(* Logix 5000 project; controller R400_500_XLS vendor 1 type 14 code 216 rev 31.11; software revision 31.01; part 27 of 32 *)
(* tags used below, declared in another part *)
   Abort1 : DINT;   // Not Used
   Alarm : SINT;   // Wait 3 seconds
   AlarmAcked : BOOL;   // Alarm has been acked
   Ashutdown : SINT;   // Not Used
   bAlrm : BOOL[64];
   Change_PrintPtr_Value : BOOL;
   CHEMICAL_COND_MAX_TIME : DINT;   // Timeout for the conductivity based chemical injection
   CHEMICAL_PUMP_OFF_TIME : DINT[4];
   CHEMICAL_PUMP_ON_TIME : DINT[4];
   CycExcBuffer : UDT_CYCLE;
   CycleSequence : UDT_CYCLE_SEQUENCE;
   CycleTime : DINT[11];   // Last cycle time saved in seconds
   DRYING : DINT;   // Drying id number
   FC23_BaseConductivity : REAL;   // Base conductivity of the water prior to the injection
   FC23_ChemicalPumpIndex : DINT;   // Chemical pump index
   FC23_CompensatedSetPoint : REAL;   // Injection compensated chemical conductivity
   FC23_FinalConductivity : REAL;   // Final value of the chemical conductivity
   FC23_OffsetSetPoint : REAL;   // Set point before enabling the on/off sequence
   FC23_ONS : SINT;
   FC23_StartSignal : BOOL;   // Conductivity based chemical injection
   FC23_WashIndex : DINT;   // Current index of the wash treatment
   FINALRINSE_1 : DINT;   // Final rinse 1 id number
   Inj_Cond : SINT;   // Conductivity injection based steps
   Inj_Cond_Tran : SINT;   // Conductivity injection based transitions
   InjMan : SINT;
   M : DINT[5];   // Memory Bits
   New_Value : SINT;
   ONS_FC24 : SINT;
   ONS_FC37 : DINT;
   ONS_FC64 : DINT;
   OPR_16_TreatPrint_Ptr : DINT;
   PREWASH_1 : DINT;   // Pre-wash 1 id number
   PREWASH_2 : DINT;   // Pre-wash 2 id number
   PREWASH_3 : DINT;   // Pre-wash 3 id number
   PREWASH_4 : DINT;   // Pre-wash 4 id number
   Print_Data : BOOL;   // Print Treatment data
   Print_Speed_Water : BOOL;
   Print_TreatEnd_Start_Data : BOOL;   // 2nd treatment of the cycle is started, pirnt Treatment Completed and Treatment data
   Print_TreatStart_Data : BOOL;   // Cycle is started Print start time and treatment data of the first treatment of the cycle
   printTreatString : STRING[85];   // Treatment String
   PWR_PrintBuffer : UDT_WASH;
   rIn_WSH61 : REAL;
   RINSE_1 : DINT;   // Rinse 1 id number
   RINSE_2 : DINT;   // Rinse 2 id number
   RINSE_3 : DINT;   // Rinse 3 id number
   RINSE_4 : DINT;   // Rinse 4 id number
   Run : DINT;
   sCRLF : STRING;
   SET_POINT_FRACTION : REAL[4];
   sFll_Zero : STRING[20];
   SMART_MODE_DRYING_HEATCOOL_SEC : DINT;   // Heating and cooling time constant for the smart mode drying (sec.)
   sOut_WSH61 : STRING;
   sPrntArray : STRING[300];   // Printer String Array
   SRE3_Serial_Number : STRING;   // Serial number
   StartPump3 : BOOL;   // Main Pump running
   String : STRING[50];   // String
   String_Temp : STRING;
   Tmr : TIMER[107];
   TreatmentPrint_Ptr : SINT;
   Trt_Drying : SINT;
   Trt_Wsh : DINT;
   VENTING : DINT;   // Venting id number
   WASH_1 : DINT;   // Wash 1 id number
   WASH_2 : DINT;   // Wash 2 id number
   WASH_3 : DINT;   // Wash 3 id number
   WASH_4 : DINT;   // Wash 4 id number
   WASH_5 : DINT;   // Wash 5 id number
   WSH36_CycleTimePercentage : DINT;
   WSH36_SecondsRemaining : DINT;
   WSH36_TotalMinutesRemaining : DINT;
   WSH36_TotalSecondsRemaining : DINT;
   WSH41_Start_signal : BOOL;   // Start cycle signal One shot rising edge
   WSH56_TreatmentInfo : BOOL;   // Treatment information for the conductivity injection
   Zero_Value : SINT;
   ChemCond : REAL;
   ChemicalName : STRING[9];   // Used by HMI
   COOLING_PHASE_TIME : DINT;   // Time of the cooling phase when time based drying
   CyclePtr : DINT;   // Cycle Pointeur
   I_Chm_1_Lvl_Sw : BOOL;   // Chemical Pump #1 level switch
   I_Chm_2_Lvl_Sw : BOOL;   // Chemical Pump #2 level switch
   I_Chm_3_Lvl_Sw : BOOL;   // Chemical Pump #3 level switch
   I_Chm_4_Lvl_Sw : BOOL;   // Chemical Pump #4 level switch
   Load : Doors;
   PrintChemCondValue : REAL;
   printID : STRING[6];
   PrintIndex : DINT;
   rSCADACompensatedSetPoint : REAL;
   Screen_Ctrl : DINT;   // PLC Screen Request
   sTime : STRING;   // String current time
   SumpTemp : REAL;   // Sump temperature in °C
   TempUnit : BOOL;   // Temperature Units 0= Celcius 1 = Farhenheit
   Tpb : DINT[11];
   TreatmentPtr : DINT;
   Unit : Hrdwre;   // Unit Configuration
(* MainProgram, continued *)

ROUTINE WSH_33_MANUAL_INJECTION   (* ladder *)
// This routine manages the manual  chemical injection
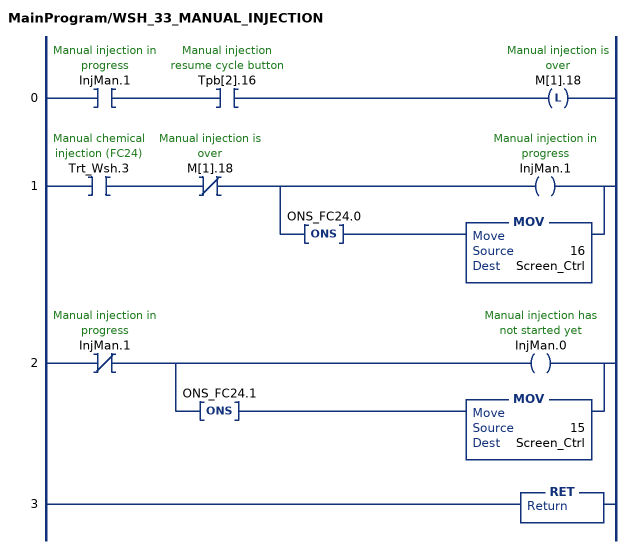
   0: XIC(InjMan.1)XIC(Tpb[2].16)OTL(M[1].18);
   1: XIC(Trt_Wsh.3)XIO(M[1].18)[OTE(InjMan.1) ,ONS(ONS_FC24.0) MOV(16,Screen_Ctrl) ];
   2: XIO(InjMan.1)[OTE(InjMan.0) ,ONS(ONS_FC24.1) MOV(15,Screen_Ctrl) ];
   3: RET();
END_ROUTINE

ROUTINE WSH_34_CONDUCTIVITY_INJECTION   (* ladder *)
// This routine manages the time based chemical injection
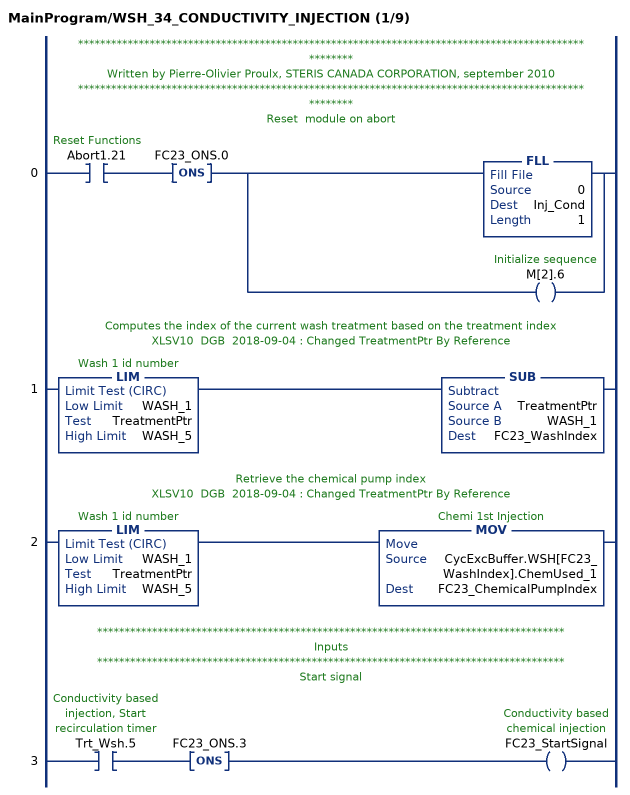
   // ****************************************************************************************************
   // Written by Pierre-Olivier Proulx, STERIS CANADA CORPORATION, september 2010
   // ****************************************************************************************************
   // Reset  module on abort
   0: XIC(Abort1.21)ONS(FC23_ONS.0)[FLL(0,Inj_Cond,1) ,OTE(M[2].6) ];
   // Computes the index of the current wash treatment based on the treatment index
   // XLSV10  DGB  2018-09-04 : Changed TreatmentPtr By Reference
   1: LIM(WASH_1,TreatmentPtr,WASH_5)SUB(TreatmentPtr,WASH_1,FC23_WashIndex);
   // Retrieve the chemical pump index
   // XLSV10  DGB  2018-09-04 : Changed TreatmentPtr By Reference
   2: LIM(WASH_1,TreatmentPtr,WASH_5)MOV(CycExcBuffer.WSH[FC23_WashIndex].ChemUsed_1,FC23_ChemicalPumpIndex);
   // *************************************************************************************
   // Inputs
   // *************************************************************************************
   // Start signal
   3: XIC(Trt_Wsh.5)ONS(FC23_ONS.3)OTE(FC23_StartSignal);
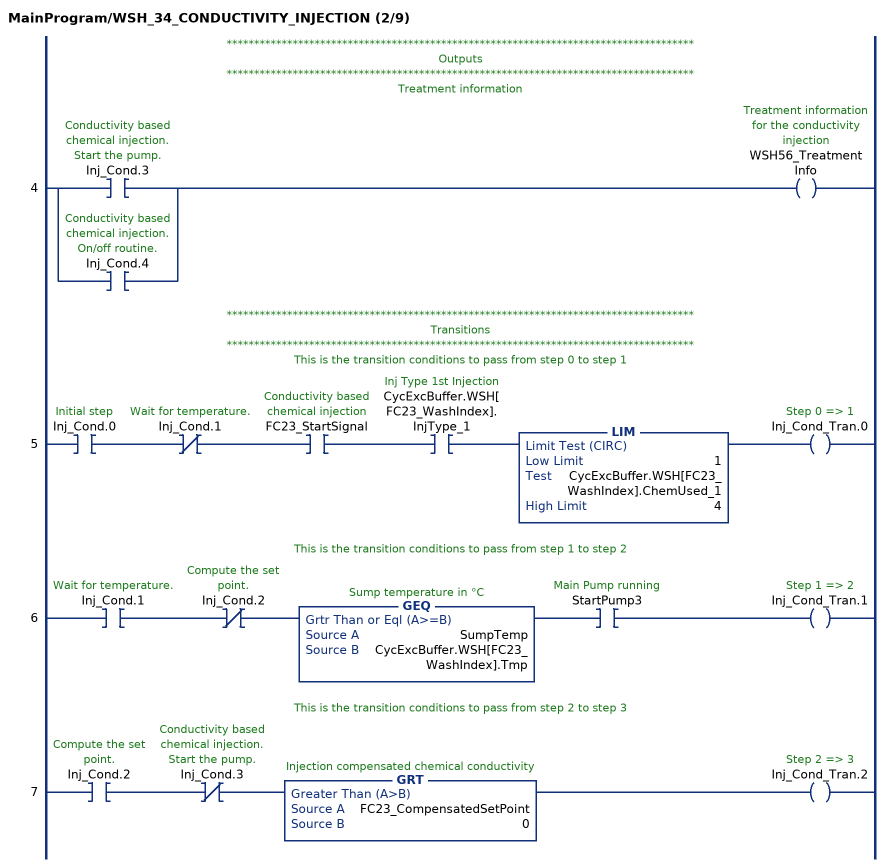
   // *************************************************************************************
   // Outputs
   // *************************************************************************************
   // Treatment information
   4: [XIC(Inj_Cond.3) ,XIC(Inj_Cond.4) ]OTE(WSH56_TreatmentInfo);
   // *************************************************************************************
   // Transitions
   // *************************************************************************************
   // This is the transition conditions to pass from step 0 to step 1
   5: XIC(Inj_Cond.0)XIO(Inj_Cond.1)XIC(FC23_StartSignal)XIC(CycExcBuffer.WSH[FC23_WashIndex].InjType_1)LIM(1,CycExcBuffer.WSH[FC23_WashIndex].ChemUsed_1,4)OTE(Inj_Cond_Tran.0);
   // This is the transition conditions to pass from step 1 to step 2
   6: XIC(Inj_Cond.1)XIO(Inj_Cond.2)GEQ(SumpTemp,CycExcBuffer.WSH[FC23_WashIndex].Tmp)XIC(StartPump3)OTE(Inj_Cond_Tran.1);
   // This is the transition conditions to pass from step 2 to step 3
   7: XIC(Inj_Cond.2)XIO(Inj_Cond.3)GRT(FC23_CompensatedSetPoint,0)OTE(Inj_Cond_Tran.2);
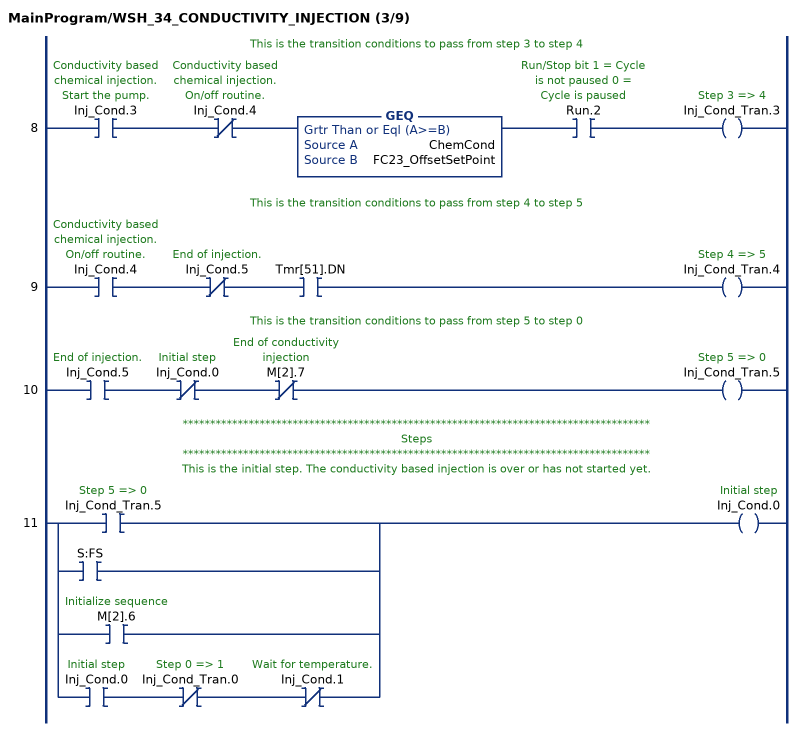
   // This is the transition conditions to pass from step 3 to step 4
   8: XIC(Inj_Cond.3)XIO(Inj_Cond.4)GEQ(ChemCond,FC23_OffsetSetPoint)XIC(Run.2)OTE(Inj_Cond_Tran.3);
   // This is the transition conditions to pass from step 4 to step 5
   9: XIC(Inj_Cond.4)XIO(Inj_Cond.5)XIC(Tmr[51].DN)OTE(Inj_Cond_Tran.4);
   // This is the transition conditions to pass from step 5 to step 0
   10: XIC(Inj_Cond.5)XIO(Inj_Cond.0)XIO(M[2].7)OTE(Inj_Cond_Tran.5);
   // *************************************************************************************
   // Steps
   // *************************************************************************************
   // This is the initial step. The conductivity based injection is over or has not started yet.
   11: [XIC(Inj_Cond_Tran.5) ,XIC(S:FS) ,XIC(M[2].6) ,XIC(Inj_Cond.0) XIO(Inj_Cond_Tran.0) XIO(Inj_Cond.1) ]OTE(Inj_Cond.0);
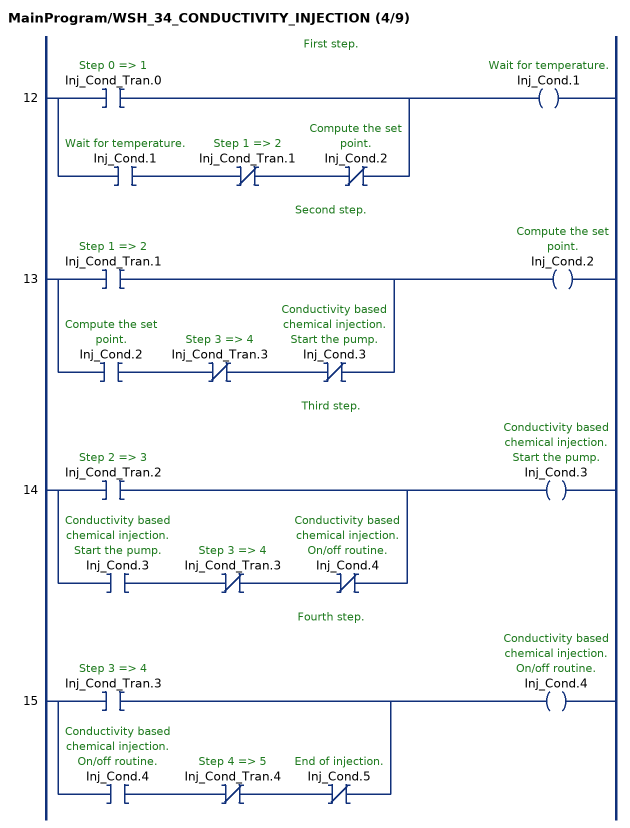
   // First step.
   12: [XIC(Inj_Cond_Tran.0) ,XIC(Inj_Cond.1) XIO(Inj_Cond_Tran.1) XIO(Inj_Cond.2) ]OTE(Inj_Cond.1);
   // Second step.
   13: [XIC(Inj_Cond_Tran.1) ,XIC(Inj_Cond.2) XIO(Inj_Cond_Tran.3) XIO(Inj_Cond.3) ]OTE(Inj_Cond.2);
   // Third step.
   14: [XIC(Inj_Cond_Tran.2) ,XIC(Inj_Cond.3) XIO(Inj_Cond_Tran.3) XIO(Inj_Cond.4) ]OTE(Inj_Cond.3);
   // Fourth step.
   15: [XIC(Inj_Cond_Tran.3) ,XIC(Inj_Cond.4) XIO(Inj_Cond_Tran.4) XIO(Inj_Cond.5) ]OTE(Inj_Cond.4);
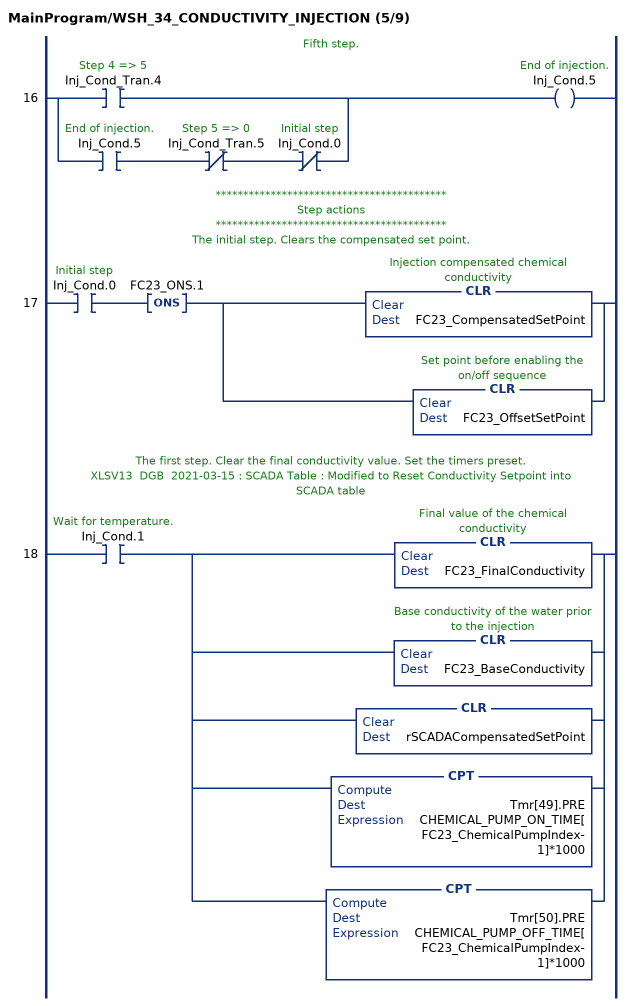
   // Fifth step.
   16: [XIC(Inj_Cond_Tran.4) ,XIC(Inj_Cond.5) XIO(Inj_Cond_Tran.5) XIO(Inj_Cond.0) ]OTE(Inj_Cond.5);
   // ******************************************
   // Step actions
   // ******************************************
   // The initial step. Clears the compensated set point.
   17: XIC(Inj_Cond.0)ONS(FC23_ONS.1)[CLR(FC23_CompensatedSetPoint) ,CLR(FC23_OffsetSetPoint) ];
   // The first step. Clear the final conductivity value. Set the timers preset.
   // XLSV13  DGB  2021-03-15 : SCADA Table : Modified to Reset Conductivity Setpoint into SCADA table
   18: XIC(Inj_Cond.1)[CLR(FC23_FinalConductivity) ,CLR(FC23_BaseConductivity) ,CLR(rSCADACompensatedSetPoint) ,CPT(Tmr[49].PRE,CHEMICAL_PUMP_ON_TIME[FC23_ChemicalPumpIndex-1]*1000) ,CPT(Tmr[50].PRE,CHEMICAL_PUMP_OFF_TIME[FC23_ChemicalPumpIndex-1]*1000) ];
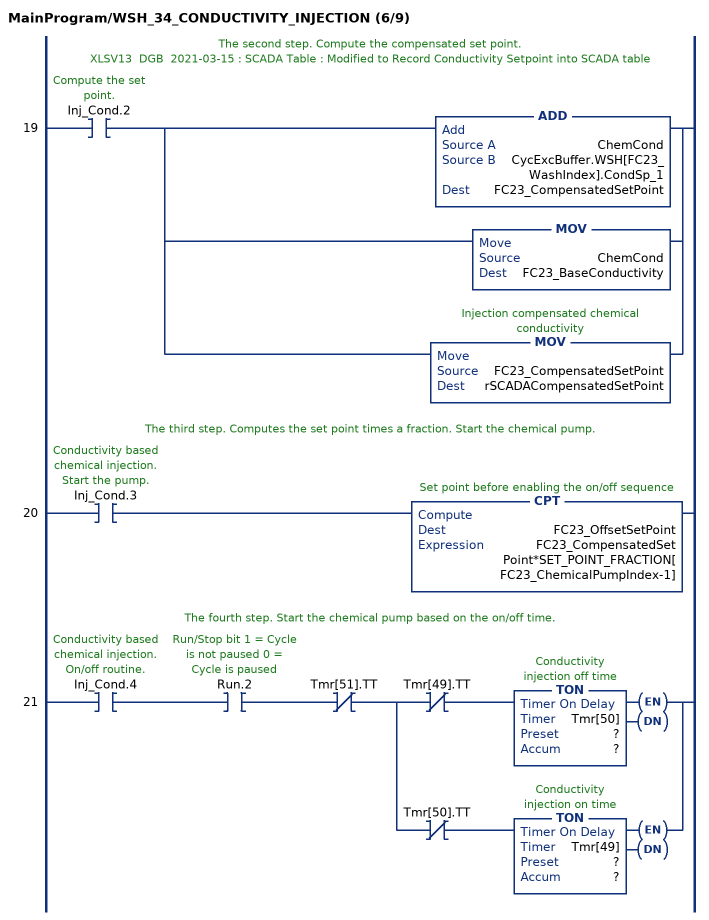
   // The second step. Compute the compensated set point.
   // XLSV13  DGB  2021-03-15 : SCADA Table : Modified to Record Conductivity Setpoint into SCADA table
   19: XIC(Inj_Cond.2)[ADD(ChemCond,CycExcBuffer.WSH[FC23_WashIndex].CondSp_1,FC23_CompensatedSetPoint) ,MOV(ChemCond,FC23_BaseConductivity) ,MOV(FC23_CompensatedSetPoint,rSCADACompensatedSetPoint) ];
   // The third step. Computes the set point times a fraction. Start the chemical pump.
   20: XIC(Inj_Cond.3)CPT(FC23_OffsetSetPoint,FC23_CompensatedSetPoint*SET_POINT_FRACTION[FC23_ChemicalPumpIndex-1]);
   // The fourth step. Start the chemical pump based on the on/off time.
   21: XIC(Inj_Cond.4)XIC(Run.2)XIO(Tmr[51].TT)[XIO(Tmr[49].TT) TON(Tmr[50],?,?) ,XIO(Tmr[50].TT) TON(Tmr[49],?,?) ];
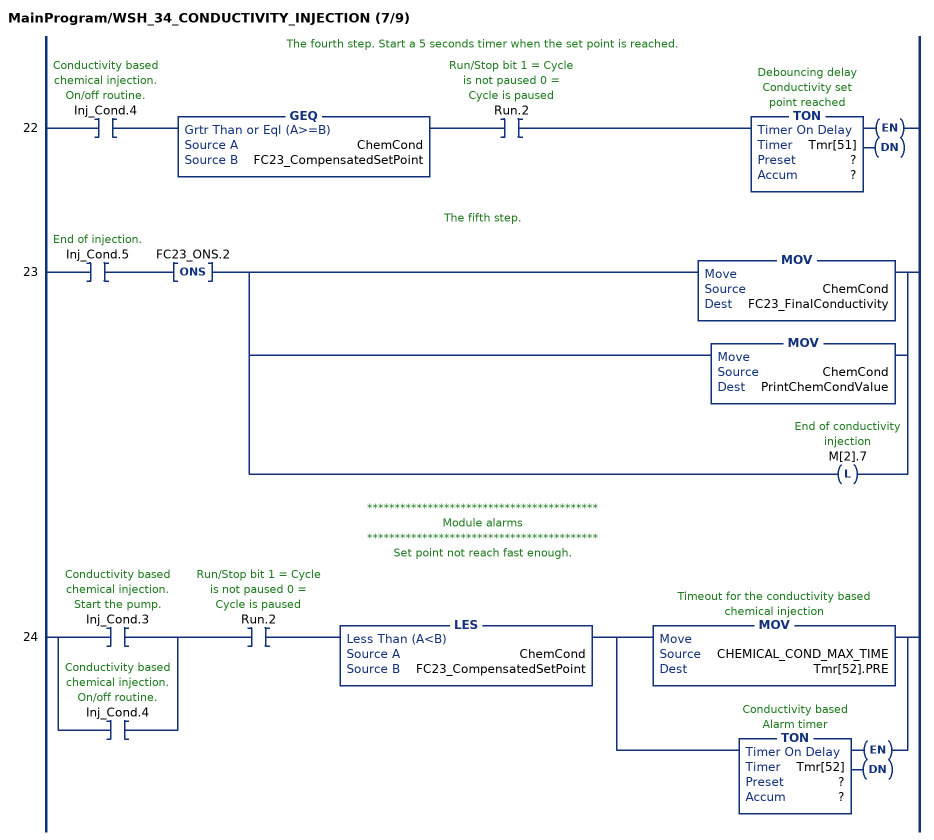
   // The fourth step. Start a 5 seconds timer when the set point is reached.
   22: XIC(Inj_Cond.4)GEQ(ChemCond,FC23_CompensatedSetPoint)XIC(Run.2)TON(Tmr[51],?,?);
   // The fifth step.
   23: XIC(Inj_Cond.5)ONS(FC23_ONS.2)[MOV(ChemCond,FC23_FinalConductivity) ,MOV(ChemCond,PrintChemCondValue) ,OTL(M[2].7) ];
   // ******************************************
   // Module alarms
   // ******************************************
   // Set point not reach fast enough.
   24: [XIC(Inj_Cond.3) ,XIC(Inj_Cond.4) ]XIC(Run.2)LES(ChemCond,FC23_CompensatedSetPoint)[MOV(CHEMICAL_COND_MAX_TIME,Tmr[52].PRE) ,TON(Tmr[52],?,?) ];
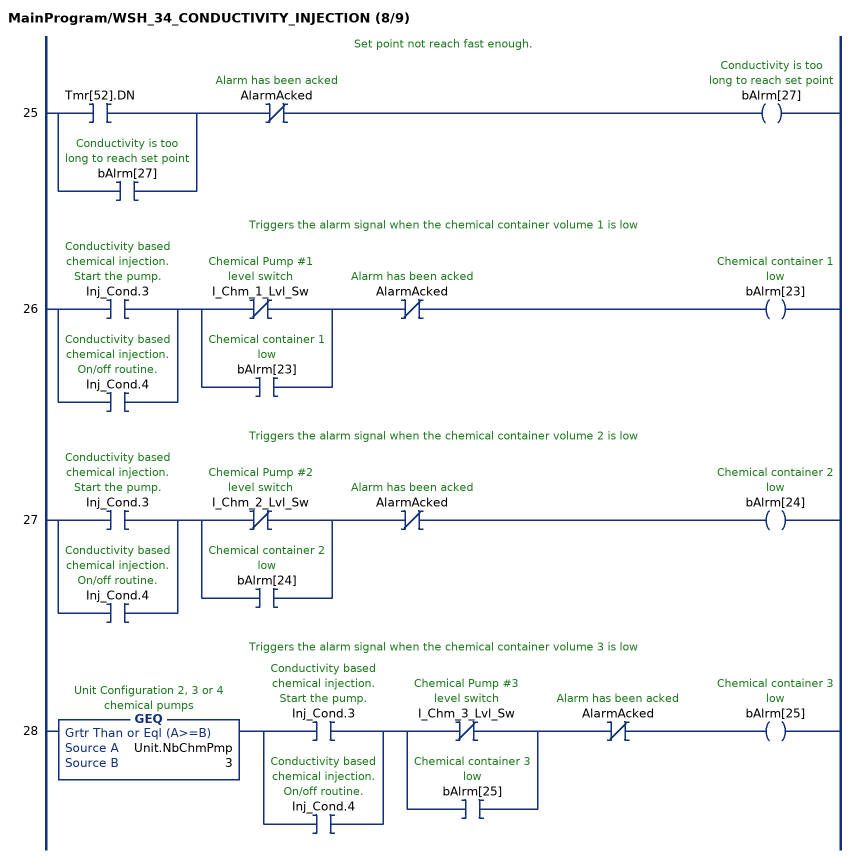
   // Set point not reach fast enough.
   25: [XIC(Tmr[52].DN) ,XIC(bAlrm[27]) ]XIO(AlarmAcked)OTE(bAlrm[27]);
   // Triggers the alarm signal when the chemical container volume 1 is low
   26: [XIC(Inj_Cond.3) ,XIC(Inj_Cond.4) ][XIO(I_Chm_1_Lvl_Sw) ,XIC(bAlrm[23]) ]XIO(AlarmAcked)OTE(bAlrm[23]);
   // Triggers the alarm signal when the chemical container volume 2 is low
   27: [XIC(Inj_Cond.3) ,XIC(Inj_Cond.4) ][XIO(I_Chm_2_Lvl_Sw) ,XIC(bAlrm[24]) ]XIO(AlarmAcked)OTE(bAlrm[24]);
   // Triggers the alarm signal when the chemical container volume 3 is low
   28: GEQ(Unit.NbChmPmp,3)[XIC(Inj_Cond.3) ,XIC(Inj_Cond.4) ][XIO(I_Chm_3_Lvl_Sw) ,XIC(bAlrm[25]) ]XIO(AlarmAcked)OTE(bAlrm[25]);
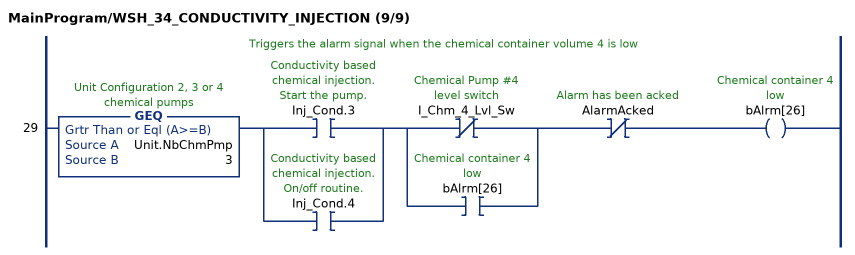
   // Triggers the alarm signal when the chemical container volume 4 is low
   29: GEQ(Unit.NbChmPmp,3)[XIC(Inj_Cond.3) ,XIC(Inj_Cond.4) ][XIO(I_Chm_4_Lvl_Sw) ,XIC(bAlrm[26]) ]XIO(AlarmAcked)OTE(bAlrm[26]);
END_ROUTINE

ROUTINE WSH_36_CycleTimeWizard   (* ladder *)
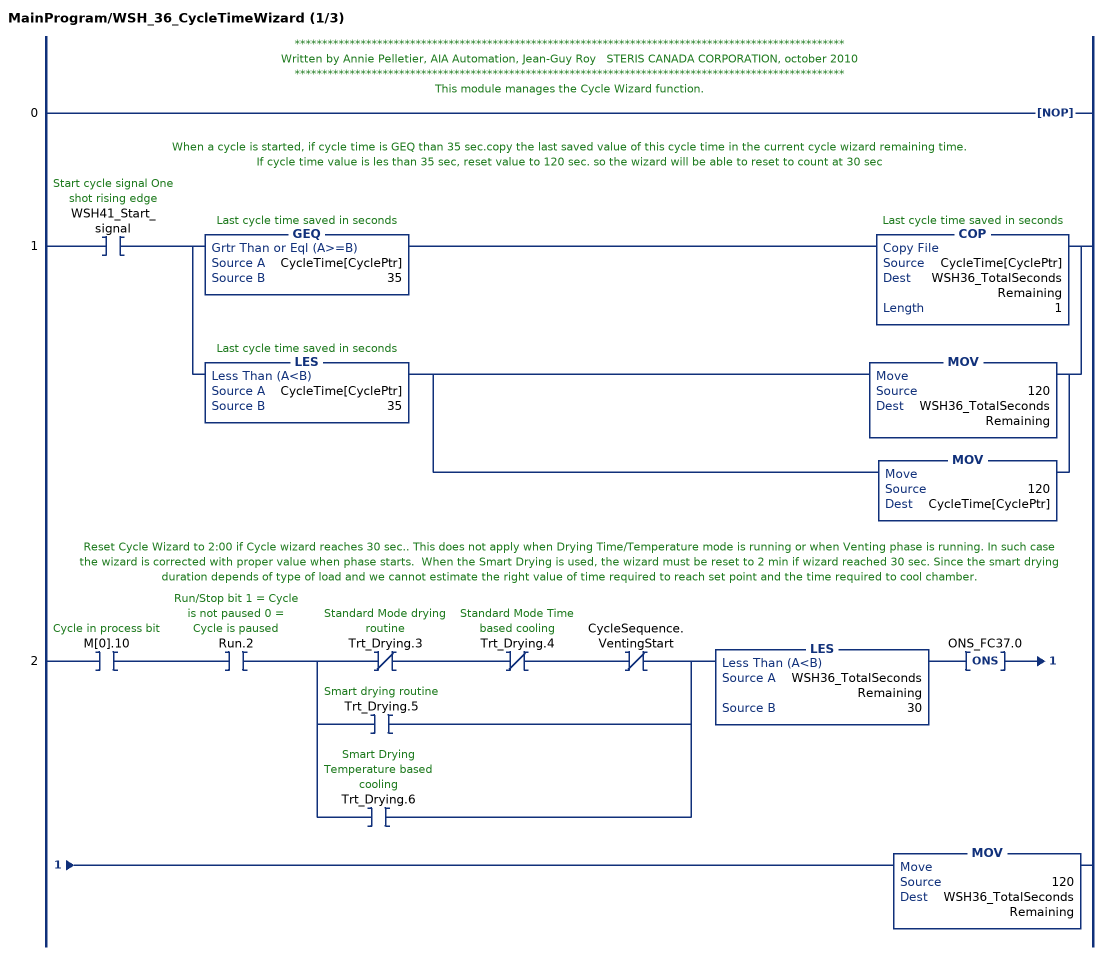
   // ****************************************************************************************************
   // Written by Annie Pelletier, AIA Automation, Jean-Guy Roy   STERIS CANADA CORPORATION, october 2010
   // ****************************************************************************************************
   // This module manages the Cycle Wizard function.
   0: NOP();
   // When a cycle is started, if cycle time is GEQ than 35 sec.copy the last saved value of this cycle time in the current cycle wizard remaining time.
   // If cycle time value is les than 35 sec, reset value to 120 sec. so the wizard will be able to reset to count at 30 sec
   1: XIC(WSH41_Start_signal)[GEQ(CycleTime[CyclePtr],35) COP(CycleTime[CyclePtr],WSH36_TotalSecondsRemaining,1) ,LES(CycleTime[CyclePtr],35) [MOV(120,WSH36_TotalSecondsRemaining) ,MOV(120,CycleTime[CyclePtr]) ] ];
   // Reset Cycle Wizard to 2:00 if Cycle wizard reaches 30 sec.. This does not apply when Drying Time/Temperature mode is running or when Venting phase is running. In such case the wizard is corrected with proper value when phase starts.  When the Smart Drying is used, the wizard must be reset to 2 min if wizard reached 30 sec. Since the smart drying duration depends of type of load and we cannot estimate the right value of time required to reach set point and the time required to cool chamber.
   2: XIC(M[0].10)XIC(Run.2)[XIO(Trt_Drying.3) XIO(Trt_Drying.4) XIO(CycleSequence.VentingStart) ,XIC(Trt_Drying.5) ,XIC(Trt_Drying.6) ]LES(WSH36_TotalSecondsRemaining,30)ONS(ONS_FC37.0)MOV(120,WSH36_TotalSecondsRemaining);
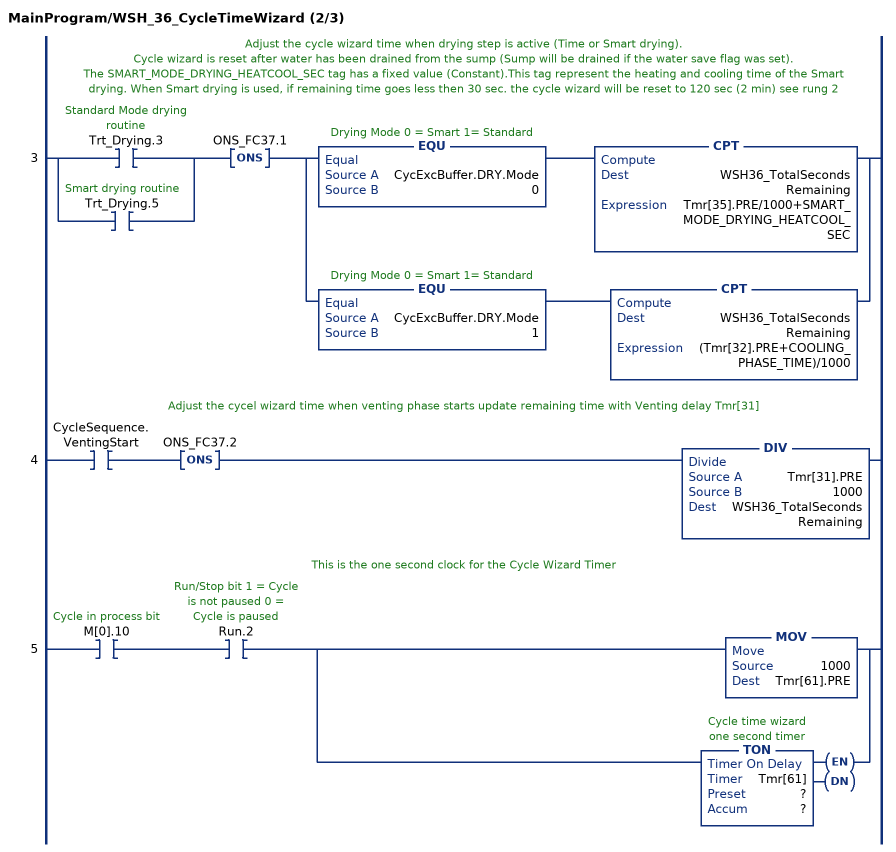
   // Adjust the cycle wizard time when drying step is active (Time or Smart drying).
   // Cycle wizard is reset after water has been drained from the sump (Sump will be drained if the water save flag was set).
   // The SMART_MODE_DRYING_HEATCOOL_SEC tag has a fixed value (Constant).This tag represent the heating and cooling time of the Smart drying. When Smart drying is used, if remaining time goes less then 30 sec. the cycle wizard will be reset to 120 sec (2 min) see rung 2
   3: [XIC(Trt_Drying.3) ,XIC(Trt_Drying.5) ]ONS(ONS_FC37.1)[EQU(CycExcBuffer.DRY.Mode,0) CPT(WSH36_TotalSecondsRemaining,Tmr[35].PRE/1000+SMART_MODE_DRYING_HEATCOOL_SEC) ,EQU(CycExcBuffer.DRY.Mode,1) CPT(WSH36_TotalSecondsRemaining,(Tmr[32].PRE+COOLING_PHASE_TIME)/1000) ];
   // Adjust the cycel wizard time when venting phase starts update remaining time with Venting delay Tmr[31]
   4: XIC(CycleSequence.VentingStart)ONS(ONS_FC37.2)DIV(Tmr[31].PRE,1000,WSH36_TotalSecondsRemaining);
   // This is the one second clock for the Cycle Wizard Timer
   5: XIC(M[0].10)XIC(Run.2)[MOV(1000,Tmr[61].PRE) ,TON(Tmr[61],?,?) ];
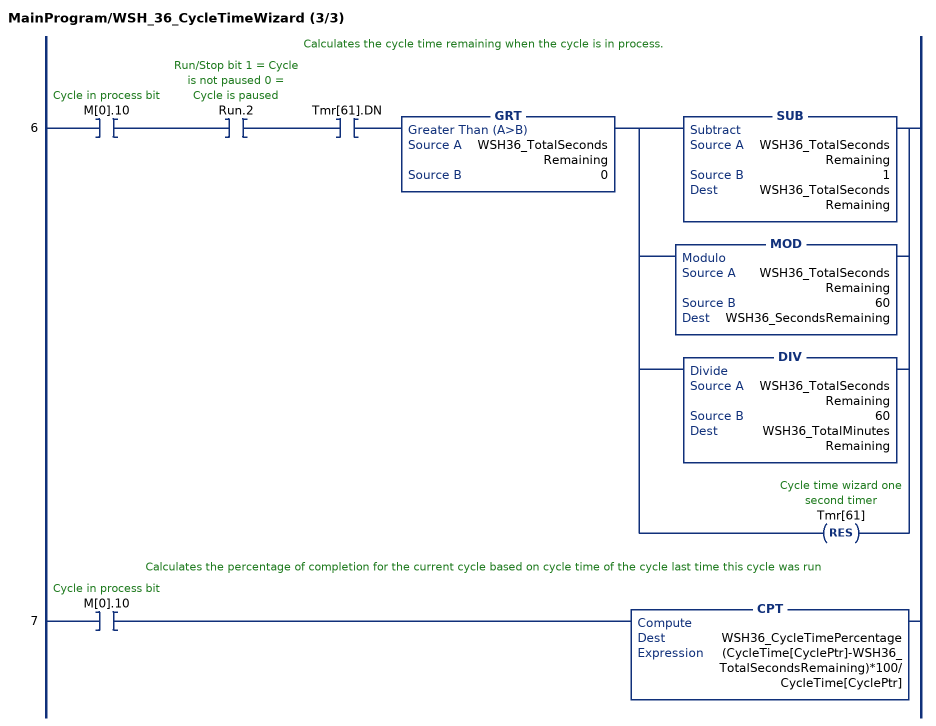
   // Calculates the cycle time remaining when the cycle is in process.
   6: XIC(M[0].10)XIC(Run.2)XIC(Tmr[61].DN)GRT(WSH36_TotalSecondsRemaining,0)[SUB(WSH36_TotalSecondsRemaining,1,WSH36_TotalSecondsRemaining) ,MOD(WSH36_TotalSecondsRemaining,60,WSH36_SecondsRemaining) ,DIV(WSH36_TotalSecondsRemaining,60,WSH36_TotalMinutesRemaining) ,RES(Tmr[61]) ];
   // Calculates the percentage of completion for the current cycle based on cycle time of the cycle last time this cycle was run
   7: XIC(M[0].10)CPT(WSH36_CycleTimePercentage,(CycleTime[CyclePtr]-WSH36_TotalSecondsRemaining)*100/CycleTime[CyclePtr]);
END_ROUTINE

ROUTINE WSH_38_GENERATE_TREAT_PAR_STRINGS   (* ladder *)
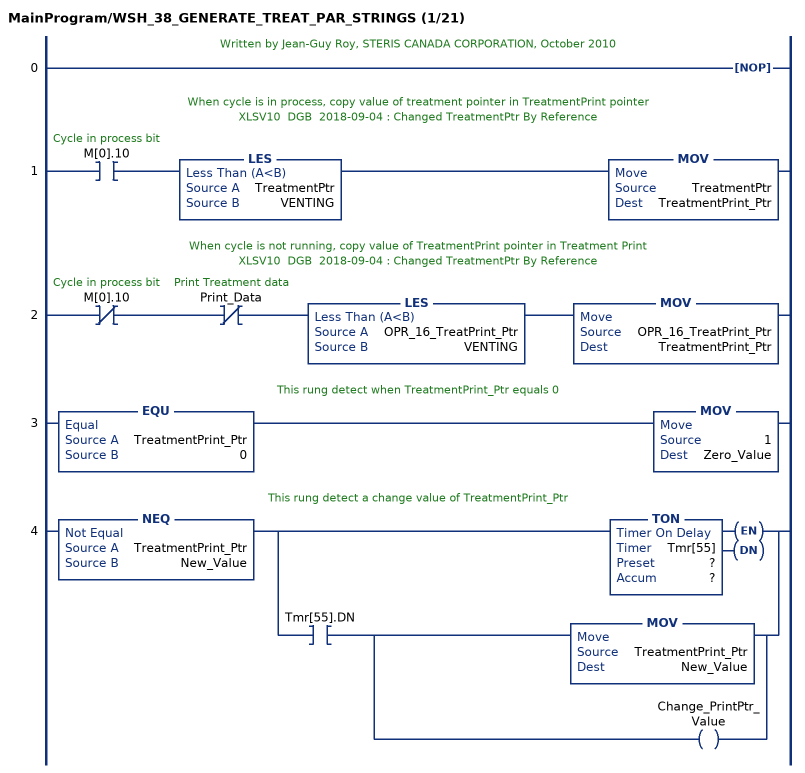
   // Written by Jean-Guy Roy, STERIS CANADA CORPORATION, October 2010
   0: NOP();
   // When cycle is in process, copy value of treatment pointer in TreatmentPrint pointer
   // XLSV10  DGB  2018-09-04 : Changed TreatmentPtr By Reference
   1: XIC(M[0].10)LES(TreatmentPtr,VENTING)MOV(TreatmentPtr,TreatmentPrint_Ptr);
   // When cycle is not running, copy value of TreatmentPrint pointer in Treatment Print
   // XLSV10  DGB  2018-09-04 : Changed TreatmentPtr By Reference
   2: XIO(M[0].10)XIO(Print_Data)LES(OPR_16_TreatPrint_Ptr,VENTING)MOV(OPR_16_TreatPrint_Ptr,TreatmentPrint_Ptr);
   // This rung detect when TreatmentPrint_Ptr equals 0
   3: EQU(TreatmentPrint_Ptr,0)MOV(1,Zero_Value);
   // This rung detect a change value of TreatmentPrint_Ptr
   4: NEQ(TreatmentPrint_Ptr,New_Value)[TON(Tmr[55],?,?) ,XIC(Tmr[55].DN) [MOV(TreatmentPrint_Ptr,New_Value) ,OTE(Change_PrintPtr_Value) ] ];
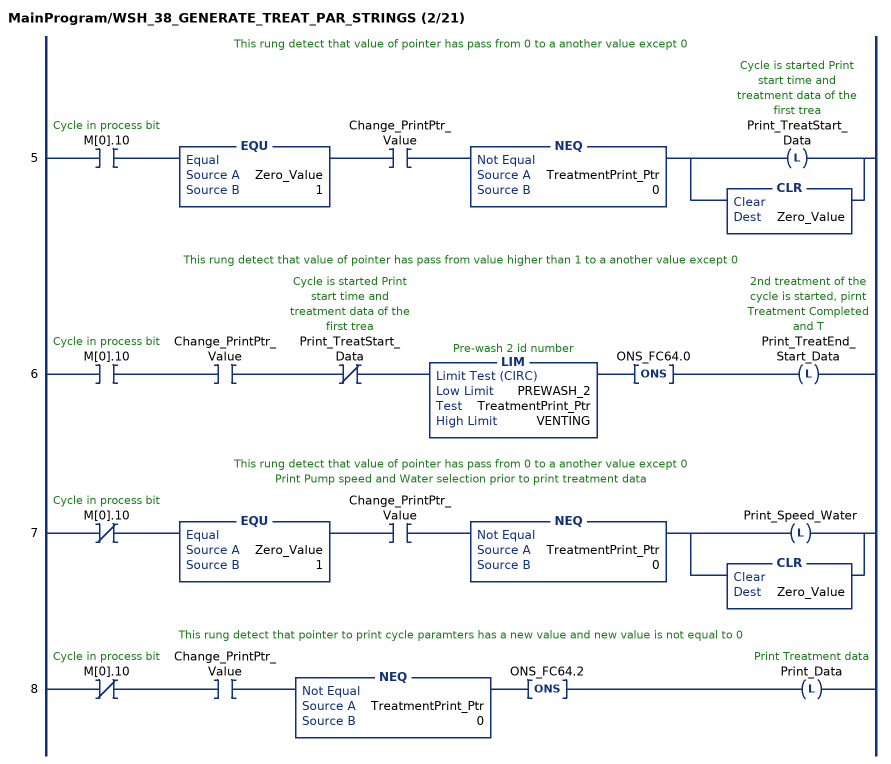
   // This rung detect that value of pointer has pass from 0 to a another value except 0
   5: XIC(M[0].10)EQU(Zero_Value,1)XIC(Change_PrintPtr_Value)NEQ(TreatmentPrint_Ptr,0)[OTL(Print_TreatStart_Data) ,CLR(Zero_Value) ];
   // This rung detect that value of pointer has pass from value higher than 1 to a another value except 0
   6: XIC(M[0].10)XIC(Change_PrintPtr_Value)XIO(Print_TreatStart_Data)LIM(PREWASH_2,TreatmentPrint_Ptr,VENTING)ONS(ONS_FC64.0)OTL(Print_TreatEnd_Start_Data);
   // This rung detect that value of pointer has pass from 0 to a another value except 0
   // Print Pump speed and Water selection prior to print treatment data
   7: XIO(M[0].10)EQU(Zero_Value,1)XIC(Change_PrintPtr_Value)NEQ(TreatmentPrint_Ptr,0)[OTL(Print_Speed_Water) ,CLR(Zero_Value) ];
   // This rung detect that pointer to print cycle paramters has a new value and new value is not equal to 0
   8: XIO(M[0].10)XIC(Change_PrintPtr_Value)NEQ(TreatmentPrint_Ptr,0)ONS(ONS_FC64.2)OTL(Print_Data);
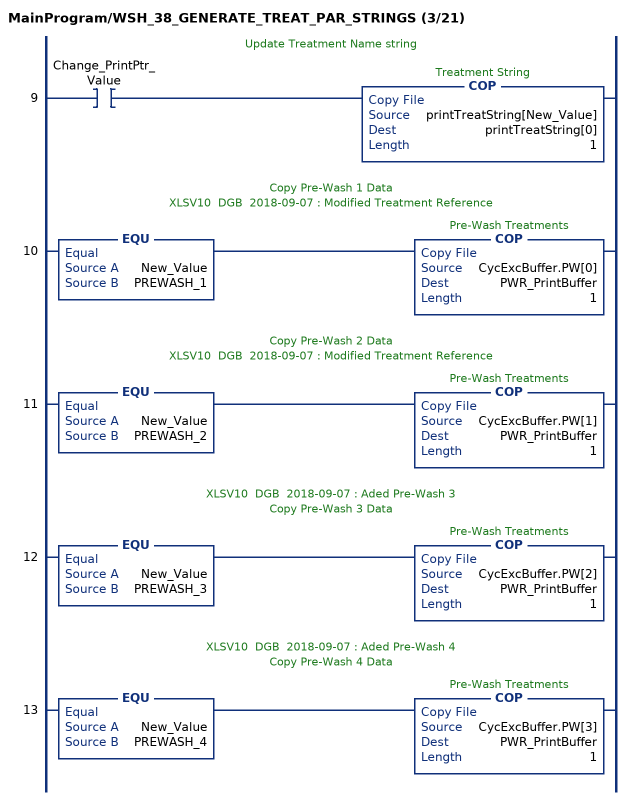
   // Update Treatment Name string
   9: XIC(Change_PrintPtr_Value)COP(printTreatString[New_Value],printTreatString[0],1);
   // Copy Pre-Wash 1 Data
   // XLSV10  DGB  2018-09-07 : Modified Treatment Reference
   10: EQU(New_Value,PREWASH_1)COP(CycExcBuffer.PW[0],PWR_PrintBuffer,1);
   // Copy Pre-Wash 2 Data
   // XLSV10  DGB  2018-09-07 : Modified Treatment Reference
   11: EQU(New_Value,PREWASH_2)COP(CycExcBuffer.PW[1],PWR_PrintBuffer,1);
   // XLSV10  DGB  2018-09-07 : Aded Pre-Wash 3
   // Copy Pre-Wash 3 Data
   12: EQU(New_Value,PREWASH_3)COP(CycExcBuffer.PW[2],PWR_PrintBuffer,1);
   // XLSV10  DGB  2018-09-07 : Aded Pre-Wash 4
   // Copy Pre-Wash 4 Data
   13: EQU(New_Value,PREWASH_4)COP(CycExcBuffer.PW[3],PWR_PrintBuffer,1);
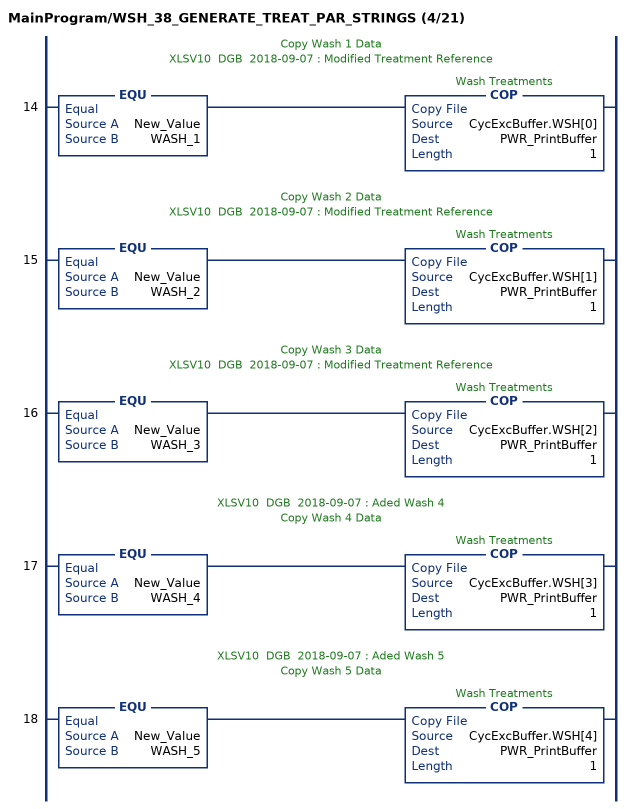
   // Copy Wash 1 Data
   // XLSV10  DGB  2018-09-07 : Modified Treatment Reference
   14: EQU(New_Value,WASH_1)COP(CycExcBuffer.WSH[0],PWR_PrintBuffer,1);
   // Copy Wash 2 Data
   // XLSV10  DGB  2018-09-07 : Modified Treatment Reference
   15: EQU(New_Value,WASH_2)COP(CycExcBuffer.WSH[1],PWR_PrintBuffer,1);
   // Copy Wash 3 Data
   // XLSV10  DGB  2018-09-07 : Modified Treatment Reference
   16: EQU(New_Value,WASH_3)COP(CycExcBuffer.WSH[2],PWR_PrintBuffer,1);
   // XLSV10  DGB  2018-09-07 : Aded Wash 4
   // Copy Wash 4 Data
   17: EQU(New_Value,WASH_4)COP(CycExcBuffer.WSH[3],PWR_PrintBuffer,1);
   // XLSV10  DGB  2018-09-07 : Aded Wash 5
   // Copy Wash 5 Data
   18: EQU(New_Value,WASH_5)COP(CycExcBuffer.WSH[4],PWR_PrintBuffer,1);
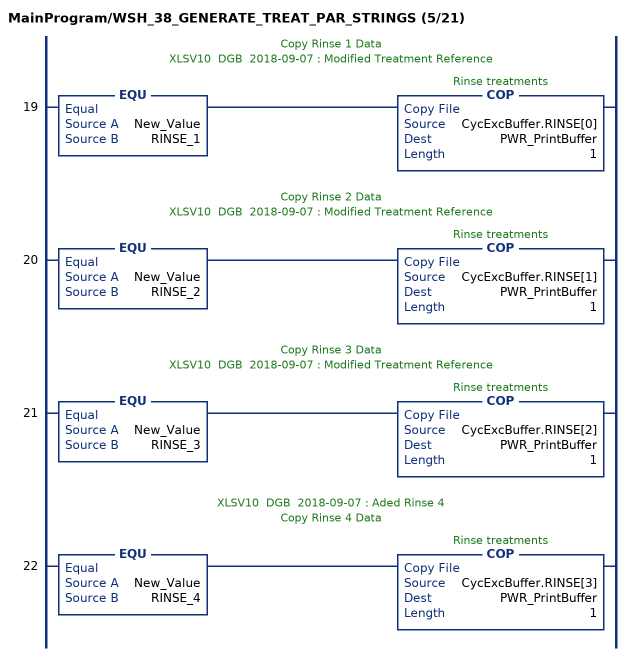
   // Copy Rinse 1 Data
   // XLSV10  DGB  2018-09-07 : Modified Treatment Reference
   19: EQU(New_Value,RINSE_1)COP(CycExcBuffer.RINSE[0],PWR_PrintBuffer,1);
   // Copy Rinse 2 Data
   // XLSV10  DGB  2018-09-07 : Modified Treatment Reference
   20: EQU(New_Value,RINSE_2)COP(CycExcBuffer.RINSE[1],PWR_PrintBuffer,1);
   // Copy Rinse 3 Data
   // XLSV10  DGB  2018-09-07 : Modified Treatment Reference
   21: EQU(New_Value,RINSE_3)COP(CycExcBuffer.RINSE[2],PWR_PrintBuffer,1);
   // XLSV10  DGB  2018-09-07 : Aded Rinse 4
   // Copy Rinse 4 Data
   22: EQU(New_Value,RINSE_4)COP(CycExcBuffer.RINSE[3],PWR_PrintBuffer,1);
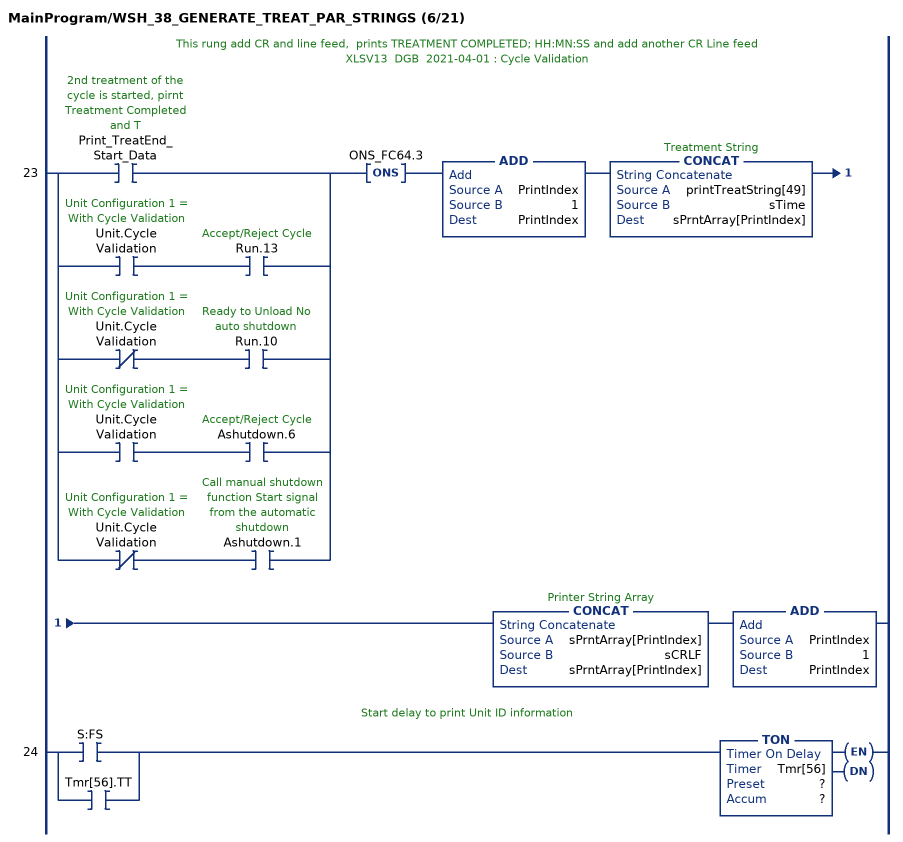
   // This rung add CR and line feed,  prints TREATMENT COMPLETED; HH:MN:SS and add another CR Line feed
   // XLSV13  DGB  2021-04-01 : Cycle Validation
   23: [XIC(Print_TreatEnd_Start_Data) ,XIC(Unit.CycleValidation) XIC(Run.13) ,XIO(Unit.CycleValidation) XIC(Run.10) ,XIC(Unit.CycleValidation) XIC(Ashutdown.6) ,XIO(Unit.CycleValidation) XIC(Ashutdown.1) ]ONS(ONS_FC64.3)ADD(PrintIndex,1,PrintIndex)CONCAT(printTreatString[49],sTime,sPrntArray[PrintIndex])CONCAT(sPrntArray[PrintIndex],sCRLF,sPrntArray[PrintIndex])ADD(PrintIndex,1,PrintIndex);
   // Start delay to print Unit ID information
   24: [XIC(S:FS) ,XIC(Tmr[56].TT) ]TON(Tmr[56],?,?);
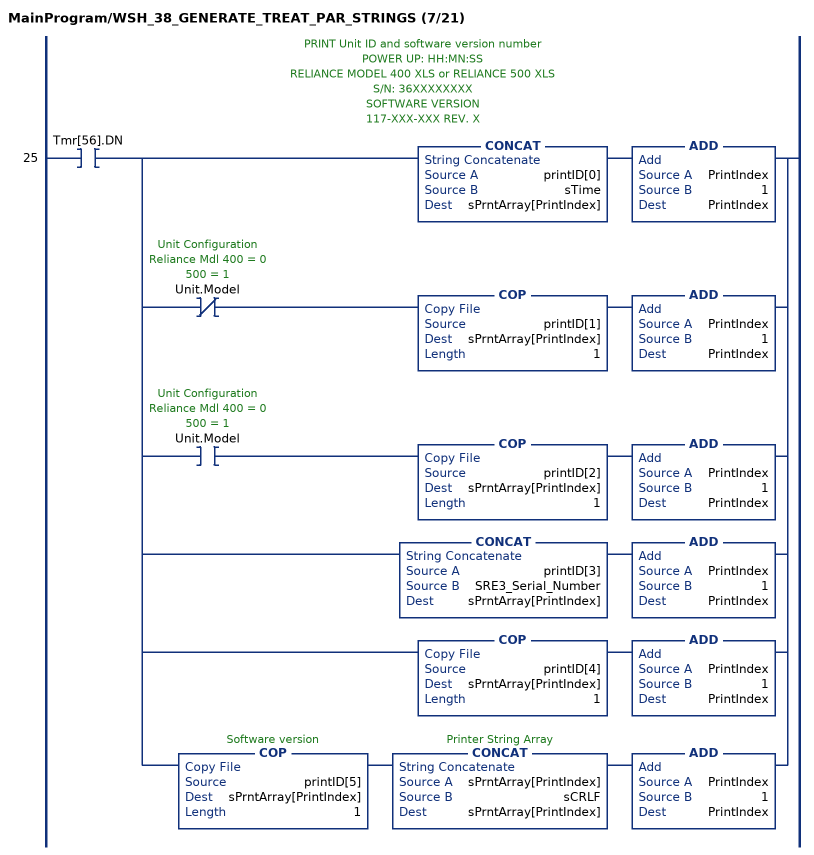
   // PRINT Unit ID and software version number
   // POWER UP: HH:MN:SS
   // RELIANCE MODEL 400 XLS or RELIANCE 500 XLS
   // S/N: 36XXXXXXXX
   // SOFTWARE VERSION
   // 117-XXX-XXX REV. X
   25: XIC(Tmr[56].DN)[CONCAT(printID[0],sTime,sPrntArray[PrintIndex]) ADD(PrintIndex,1,PrintIndex) ,XIO(Unit.Model) COP(printID[1],sPrntArray[PrintIndex],1) ADD(PrintIndex,1,PrintIndex) ,XIC(Unit.Model) COP(printID[2],sPrntArray[PrintIndex],1) ADD(PrintIndex,1,PrintIndex) ,CONCAT(printID[3],SRE3_Serial_Number,sPrntArray[PrintIndex]) ADD(PrintIndex,1,PrintIndex) ,COP(printID[4],sPrntArray[PrintIndex],1) ADD(PrintIndex,1,PrintIndex) ,COP(printID[5],sPrntArray[PrintIndex],1) CONCAT(sPrntArray[PrintIndex],sCRLF,sPrntArray[PrintIndex]) ADD(PrintIndex,1,PrintIndex) ];
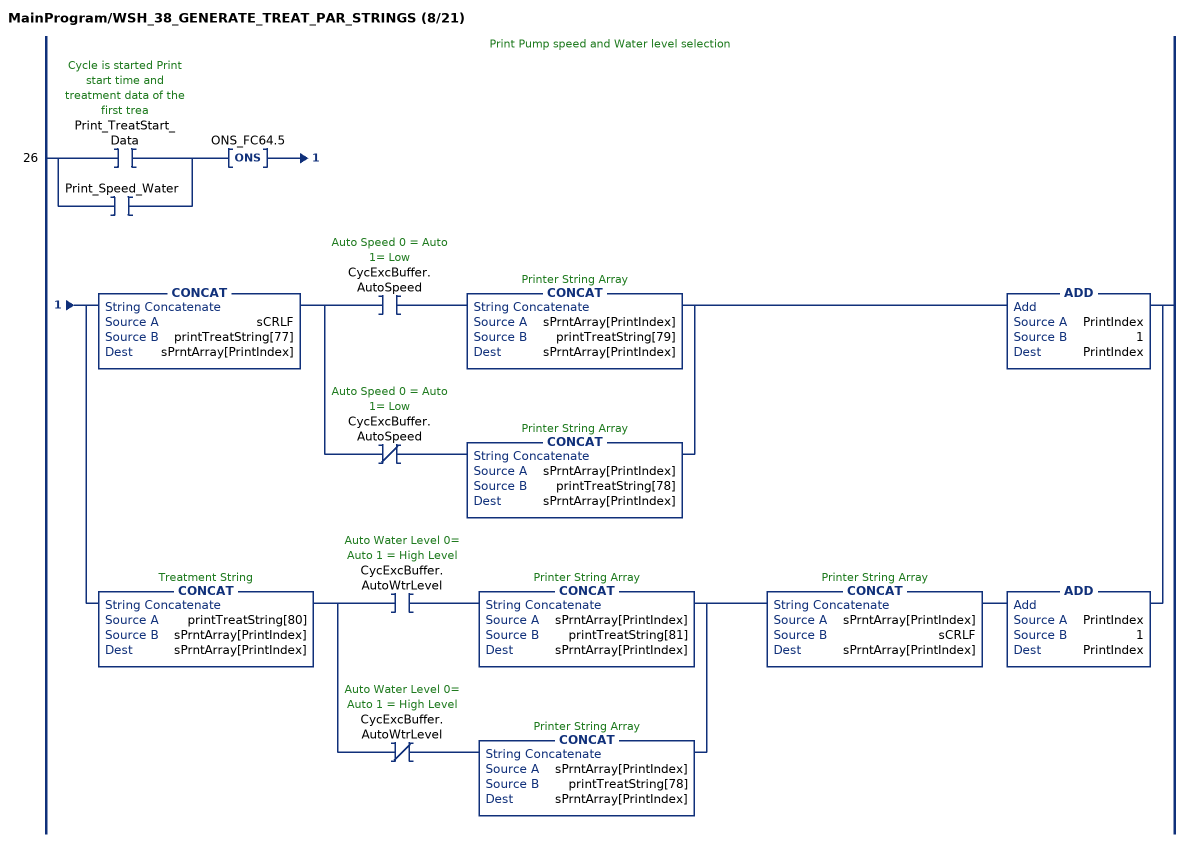
   // Print Pump speed and Water level selection
   26: [XIC(Print_TreatStart_Data) ,XIC(Print_Speed_Water) ]ONS(ONS_FC64.5)[CONCAT(sCRLF,printTreatString[77],sPrntArray[PrintIndex]) [XIC(CycExcBuffer.AutoSpeed) CONCAT(sPrntArray[PrintIndex],printTreatString[79],sPrntArray[PrintIndex]) ,XIO(CycExcBuffer.AutoSpeed) CONCAT(sPrntArray[PrintIndex],printTreatString[78],sPrntArray[PrintIndex]) ] ADD(PrintIndex,1,PrintIndex) ,CONCAT(printTreatString[80],sPrntArray[PrintIndex],sPrntArray[PrintIndex]) [XIC(CycExcBuffer.AutoWtrLevel) CONCAT(sPrntArray[PrintIndex],printTreatString[81],sPrntArray[PrintIndex]) ,XIO(CycExcBuffer.AutoWtrLevel) CONCAT(sPrntArray[PrintIndex],printTreatString[78],sPrntArray[PrintIndex]) ] CONCAT(sPrntArray[PrintIndex],sCRLF,sPrntArray[PrintIndex]) ADD(PrintIndex,1,PrintIndex) ];
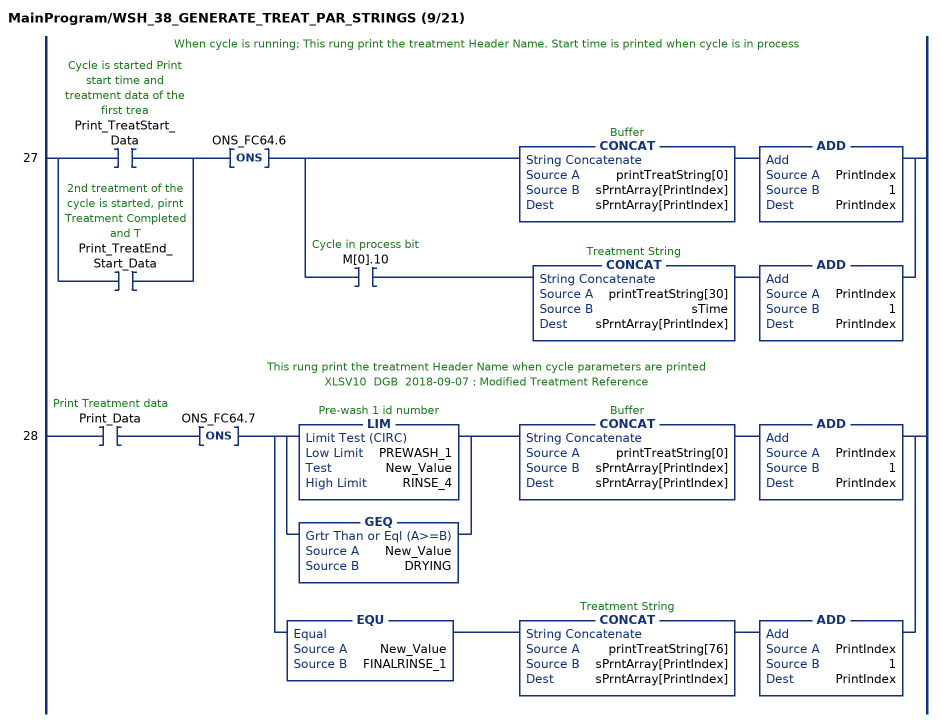
   // When cycle is running; This rung print the treatment Header Name. Start time is printed when cycle is in process
   27: [XIC(Print_TreatStart_Data) ,XIC(Print_TreatEnd_Start_Data) ]ONS(ONS_FC64.6)[CONCAT(printTreatString[0],sPrntArray[PrintIndex],sPrntArray[PrintIndex]) ADD(PrintIndex,1,PrintIndex) ,XIC(M[0].10) CONCAT(printTreatString[30],sTime,sPrntArray[PrintIndex]) ADD(PrintIndex,1,PrintIndex) ];
   // This rung print the treatment Header Name when cycle parameters are printed
   // XLSV10  DGB  2018-09-07 : Modified Treatment Reference
   28: XIC(Print_Data)ONS(ONS_FC64.7)[[LIM(PREWASH_1,New_Value,RINSE_4) ,GEQ(New_Value,DRYING) ] CONCAT(printTreatString[0],sPrntArray[PrintIndex],sPrntArray[PrintIndex]) ADD(PrintIndex,1,PrintIndex) ,EQU(New_Value,FINALRINSE_1) CONCAT(printTreatString[76],sPrntArray[PrintIndex],sPrntArray[PrintIndex]) ADD(PrintIndex,1,PrintIndex) ];
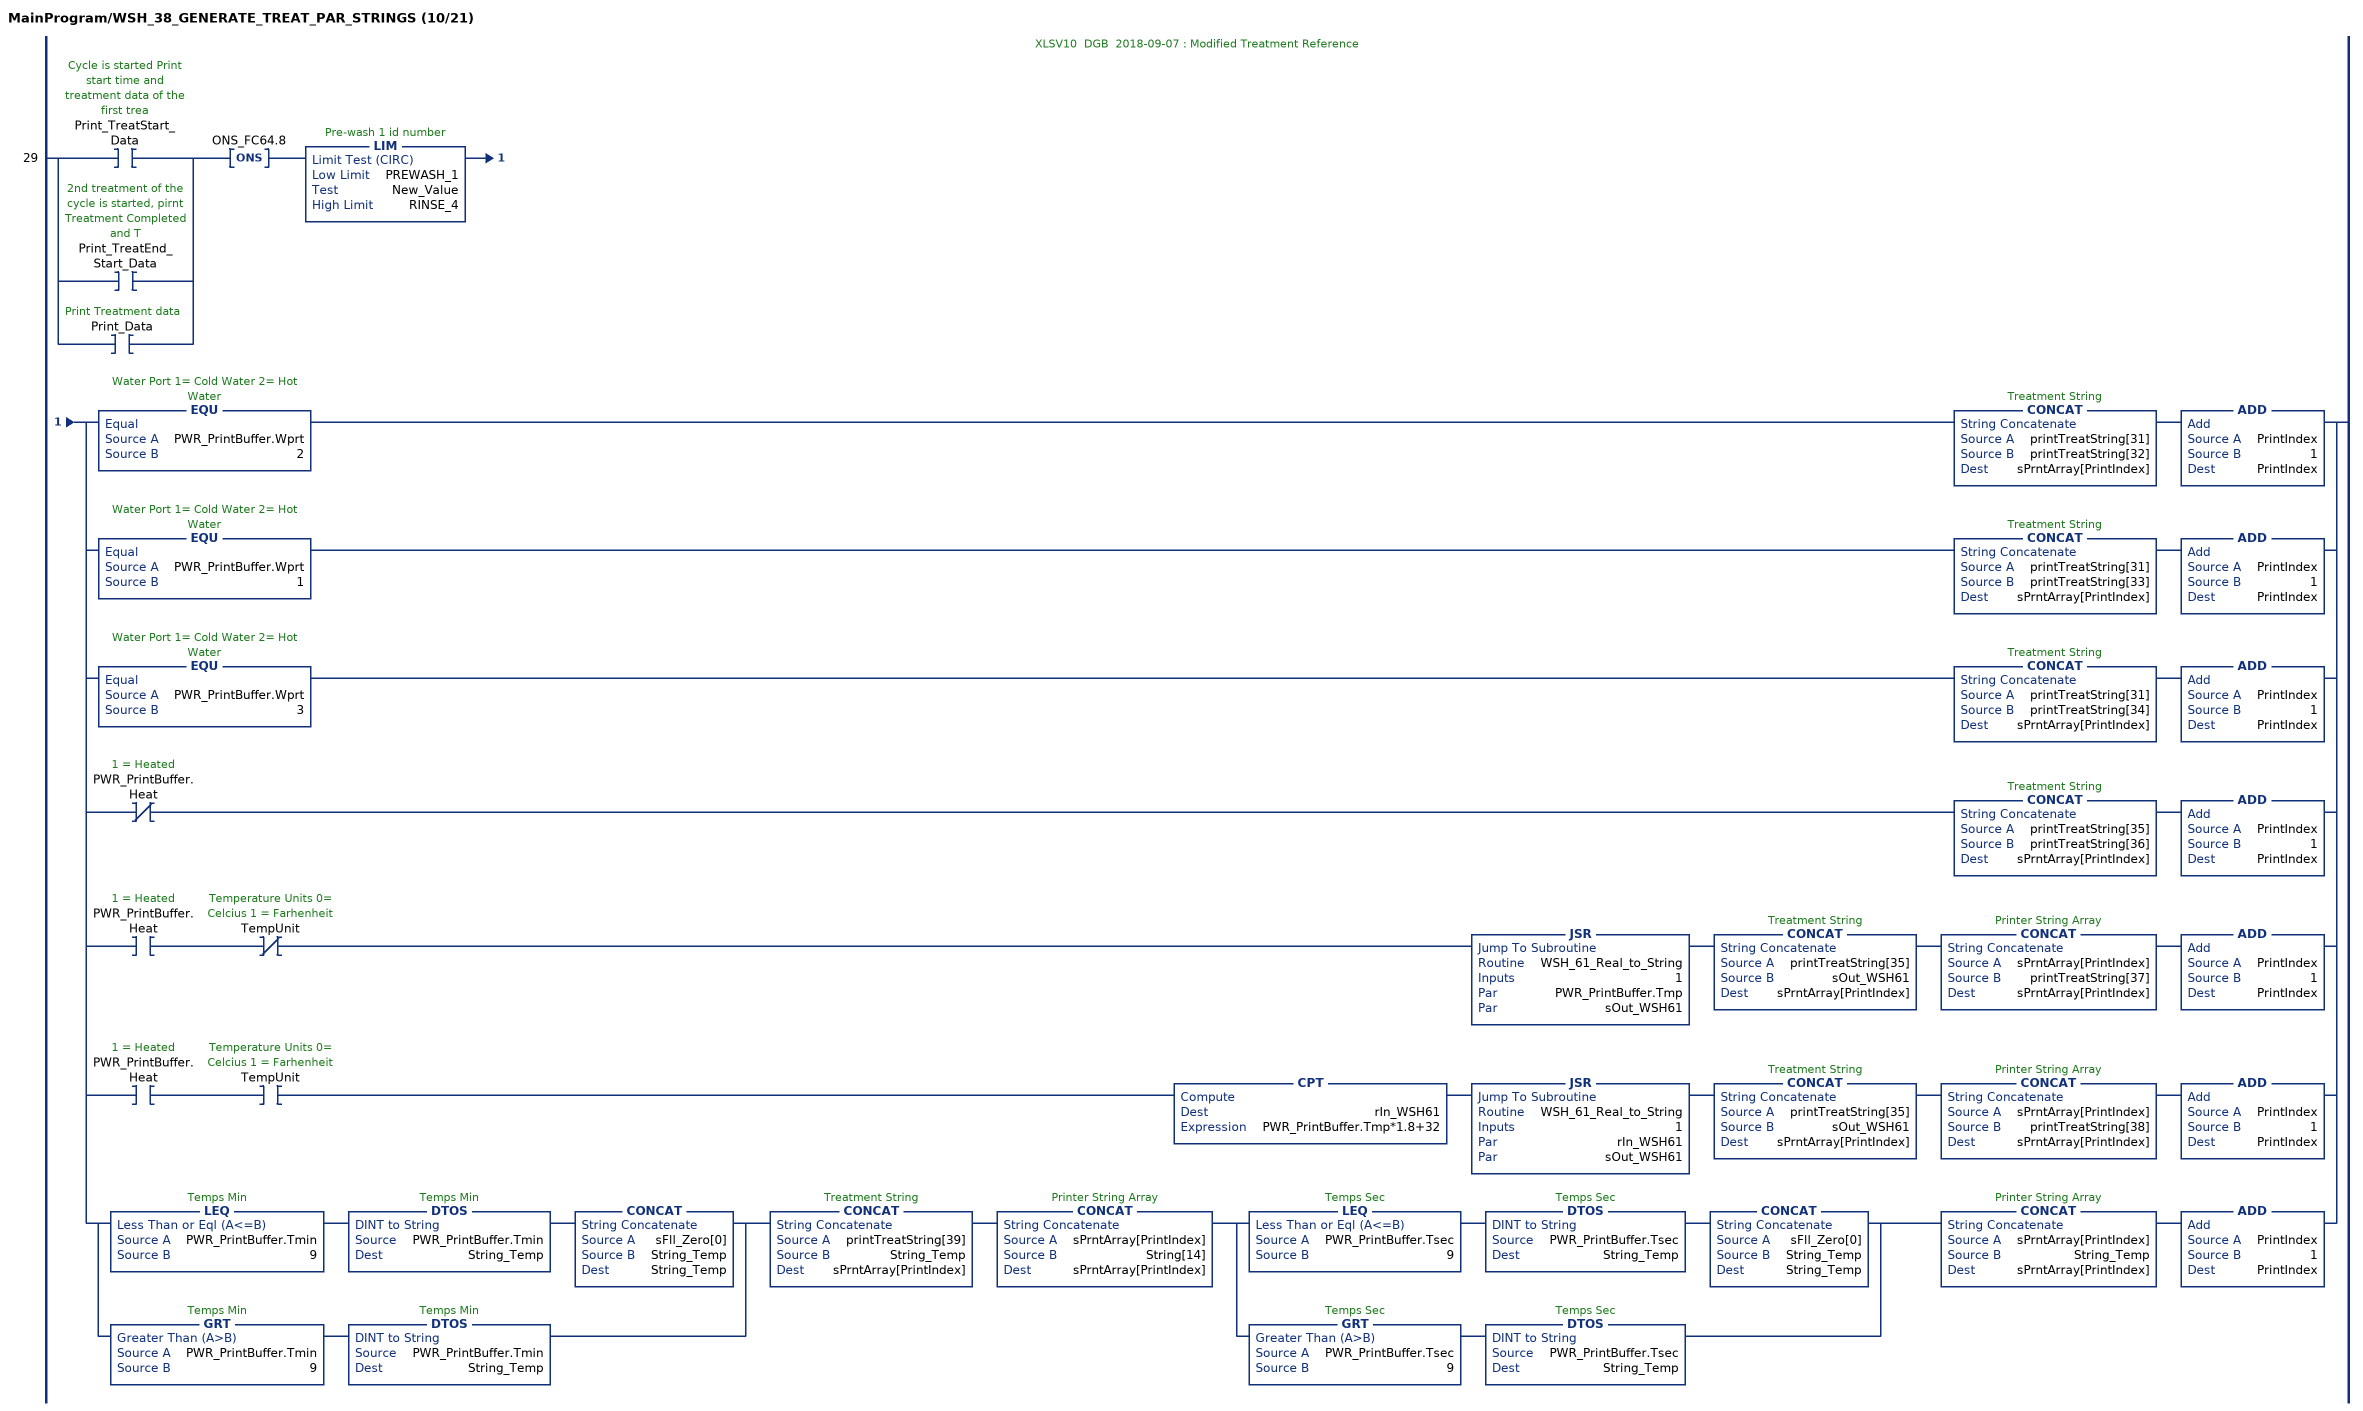
   // XLSV10  DGB  2018-09-07 : Modified Treatment Reference
   29: [XIC(Print_TreatStart_Data) ,XIC(Print_TreatEnd_Start_Data) ,XIC(Print_Data) ]ONS(ONS_FC64.8)LIM(PREWASH_1,New_Value,RINSE_4)[EQU(PWR_PrintBuffer.Wprt,2) CONCAT(printTreatString[31],printTreatString[32],sPrntArray[PrintIndex]) ADD(PrintIndex,1,PrintIndex) ,EQU(PWR_PrintBuffer.Wprt,1) CONCAT(printTreatString[31],printTreatString[33],sPrntArray[PrintIndex]) ADD(PrintIndex,1,PrintIndex) ,EQU(PWR_PrintBuffer.Wprt,3) CONCAT(printTreatString[31],printTreatString[34],sPrntArray[PrintIndex]) ADD(PrintIndex,1,PrintIndex) ,XIO(PWR_PrintBuffer.Heat) CONCAT(printTreatString[35],printTreatString[36],sPrntArray[PrintIndex]) ADD(PrintIndex,1,PrintIndex) ,XIC(PWR_PrintBuffer.Heat) XIO(TempUnit) JSR(WSH_61_Real_to_String,1,PWR_PrintBuffer.Tmp,sOut_WSH61) CONCAT(printTreatString[35],sOut_WSH61,sPrntArray[PrintIndex]) CONCAT(sPrntArray[PrintIndex],printTreatString[37],sPrntArray[PrintIndex]) ADD(PrintIndex,1,PrintIndex) ,XIC(PWR_PrintBuffer.Heat) XIC(TempUnit) CPT(rIn_WSH61,PWR_PrintBuffer.Tmp*1.8+32) JSR(WSH_61_Real_to_String,1,rIn_WSH61,sOut_WSH61) CONCAT(printTreatString[35],sOut_WSH61,sPrntArray[PrintIndex]) CONCAT(sPrntArray[PrintIndex],printTreatString[38],sPrntArray[PrintIndex]) ADD(PrintIndex,1,PrintIndex) ,[LEQ(PWR_PrintBuffer.Tmin,9) DTOS(PWR_PrintBuffer.Tmin,String_Temp) CONCAT(sFll_Zero[0],String_Temp,String_Temp) ,GRT(PWR_PrintBuffer.Tmin,9) DTOS(PWR_PrintBuffer.Tmin,String_Temp) ] CONCAT(printTreatString[39],String_Temp,sPrntArray[PrintIndex]) CONCAT(sPrntArray[PrintIndex],String[14],sPrntArray[PrintIndex]) [LEQ(PWR_PrintBuffer.Tsec,9) DTOS(PWR_PrintBuffer.Tsec,String_Temp) CONCAT(sFll_Zero[0],String_Temp,String_Temp) ,GRT(PWR_PrintBuffer.Tsec,9) DTOS(PWR_PrintBuffer.Tsec,String_Temp) ] CONCAT(sPrntArray[PrintIndex],String_Temp,sPrntArray[PrintIndex]) ADD(PrintIndex,1,PrintIndex) ];
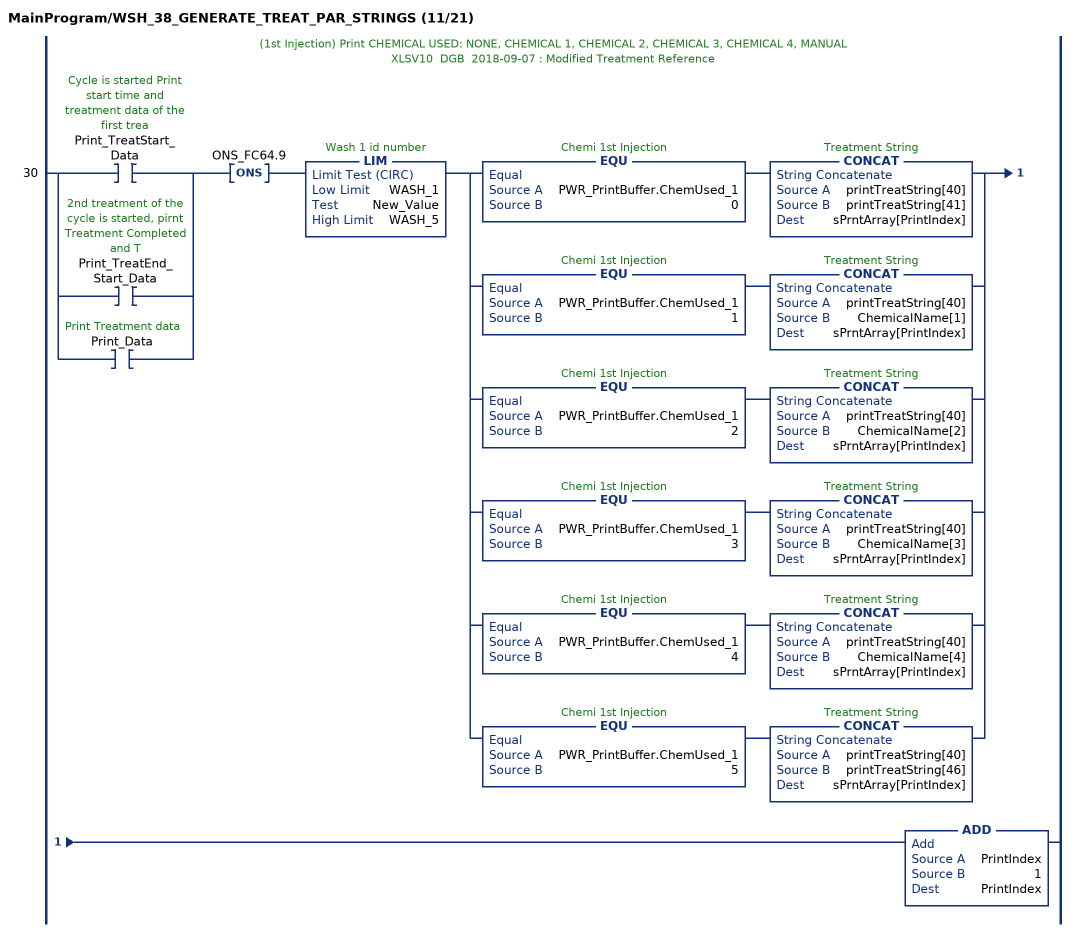
   // (1st Injection) Print CHEMICAL USED: NONE, CHEMICAL 1, CHEMICAL 2, CHEMICAL 3, CHEMICAL 4, MANUAL
   // XLSV10  DGB  2018-09-07 : Modified Treatment Reference
   30: [XIC(Print_TreatStart_Data) ,XIC(Print_TreatEnd_Start_Data) ,XIC(Print_Data) ]ONS(ONS_FC64.9)LIM(WASH_1,New_Value,WASH_5)[EQU(PWR_PrintBuffer.ChemUsed_1,0) CONCAT(printTreatString[40],printTreatString[41],sPrntArray[PrintIndex]) ,EQU(PWR_PrintBuffer.ChemUsed_1,1) CONCAT(printTreatString[40],ChemicalName[1],sPrntArray[PrintIndex]) ,EQU(PWR_PrintBuffer.ChemUsed_1,2) CONCAT(printTreatString[40],ChemicalName[2],sPrntArray[PrintIndex]) ,EQU(PWR_PrintBuffer.ChemUsed_1,3) CONCAT(printTreatString[40],ChemicalName[3],sPrntArray[PrintIndex]) ,EQU(PWR_PrintBuffer.ChemUsed_1,4) CONCAT(printTreatString[40],ChemicalName[4],sPrntArray[PrintIndex]) ,EQU(PWR_PrintBuffer.ChemUsed_1,5) CONCAT(printTreatString[40],printTreatString[46],sPrntArray[PrintIndex]) ]ADD(PrintIndex,1,PrintIndex);
